FUNCTION_BLOCK SC_MoveNeedleDown (* The contract of a skill primitive, the only part that is its own: which command it sends (and with what argument, and which when it ends), how long it may run, and three conditions on the equipment's signals and its parameters: when it may start, when it is done, what must hold while it runs. Technical: MoveNeedleDown: Precondition NOT (AtTop AND AtBottom); NeedleAxis.Down until (Position >= Distance) OR AtBottom; Invariant NOT (AtTop AND AtBottom) *)
  (* Standard: 61499-2 *)
  (* Version 0.1, 2026-09-28, Project contributors, AAU Smart Production Lab *)
  PACKAGE filler;
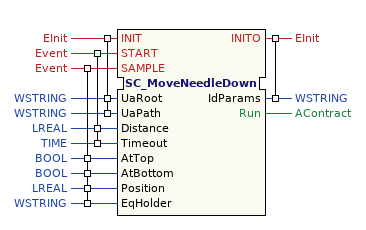
  EVENT_INPUT
    INIT : EInit WITH UaRoot, UaPath; (* Initialise: name the OPC UA variables of the parameters and results *)
    START WITH Distance, Timeout; (* A run starts, with the parameters: say what the skill does *)
    SAMPLE WITH AtTop, AtBottom, Position, EqHolder; (* The equipment's newest state arrived *)
  END_EVENT
  EVENT_OUTPUT
    INITO : EInit WITH IdParams; (* Initialised: the next block of the INIT chain goes on *)
  END_EVENT
  VAR_INPUT
    UaRoot : WSTRING; (* The module's OPC UA folder, e.g. /Objects/Filling *)
    UaPath : WSTRING; (* This skill's OPC UA folder below UaRoot, e.g. /Skills/Dispensing *)
    Distance : LREAL; (* Parameter Distance mm, 0.0 to 50.0: Target depth below the top position *)
    Timeout : TIME; (* How long the run may take before it fails with Timeout (3) *)
    AtTop : BOOL; (* NeedleAxis: AtTop, an input *)
    AtBottom : BOOL; (* NeedleAxis: AtBottom, an input *)
    Position : LREAL; (* NeedleAxis: Position (mm), an input *)
    EqHolder : WSTRING; (* Who holds the equipment now (empty: free), passed on to the run *)
  END_VAR
  VAR_OUTPUT
    IdParams : WSTRING; (* OPC UA ID of the published parameters *)
  END_VAR
  PLUGS
    Run : modlib::AContract; (* To the run (AContract): what the skill does and when it is done *)
  END_PLUGS
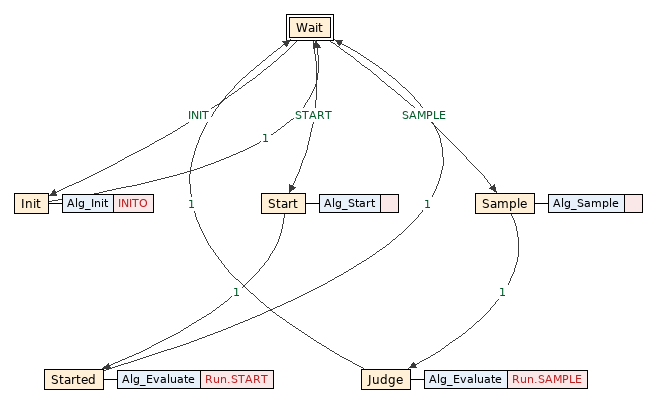
  EC_STATES
    Wait;
    Init : Alg_Init -> INITO;
    Start : Alg_Start;
    Started : Alg_Evaluate -> Run.START;
    Sample : Alg_Sample;
    Judge : Alg_Evaluate -> Run.SAMPLE;
  END_STATES
  EC_TRANSITIONS
    Wait TO Init := INIT;
    Init TO Wait := 1;
    Wait TO Start := START;
    Start TO Started := 1;
    Started TO Wait := 1;
    Wait TO Sample := SAMPLE;
    Sample TO Judge := 1;
    Judge TO Wait := 1;
  END_TRANSITIONS
  ALGORITHM Alg_Init IN ST:
IdParams := CONCAT(CONCAT(CONCAT("opc_ua[WRITE;", CONCAT(UaRoot, UaPath)), "/Parameters/Distance"), "]");
  END_ALGORITHM
  ALGORITHM Alg_Start IN ST:
Run.Timed := FALSE;
Run.RunTime := Timeout;
Run.Command := 1;
Run.Arg := 0.0;
Run.StopCommand := 0;
  END_ALGORITHM
  ALGORITHM Alg_Evaluate IN ST:
Run.Pre := NOT (AtTop AND AtBottom);
Run.Post := (Position >= Distance) OR AtBottom;
Run.Inv := NOT (AtTop AND AtBottom);
  END_ALGORITHM
  ALGORITHM Alg_Sample IN ST:
Run.EqHolder := EqHolder;
  END_ALGORITHM
END_FUNCTION_BLOCK
